TYPE ST_MasterParam :
STRUCT
	fStartPos: LREAL;
	fEndPos: LREAL;
	fVelocity: LREAL;
END_STRUCT
END_TYPE

(* stored: Version 1.1.0.1, ProductVersion 3.1.4024.12
   DUT ST_MasterParam: Id {39a2e362-02e7-48fb-aba4-245804338adc} *)
